Fanuc KAREL source: kb00188.KL

-- PROVISIONAL review KL for V940-1; original PC SHA256 6403144fd7e4112def682653404230262cf418242f487b0eccd2e369bb4e620a
-- Incomplete behavior may be omitted. Consult companion uncertainty JSON. Do not deploy.
PROGRAM KB00188
%NOLOCKGROUP
VAR
  P1 : STRING[80]
  RESULT : INTEGER
BEGIN
  -- V9_ZERO_TABLE_METADATA_HINT layout=0001; no indexed target words; source/name/runtime held
  -- UNRESOLVED_PC offsets 5-14; opcodes 3F,75
  -- UNRESOLVED_PC offsets 19-36; opcodes 27,22,2A,76,23
  -- UNRESOLVED_PC offsets 41-45; opcodes 7F
END KB00188
